FUNCTION_BLOCK R2 (* Basic Function Block Type *)
  (* Standard: 61499-2 *)
  (* Version 0.0, 10/11/2026, lizar, nxtControl GmBH, Template *)
  PACKAGE Main;
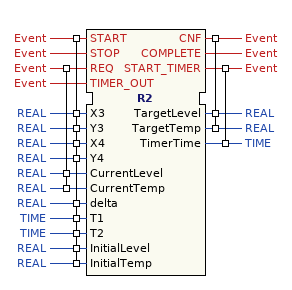
  EVENT_INPUT
    START WITH X3, Y3, X4, Y4, delta, T1, T2, InitialLevel, InitialTemp; (* Normal Execution Request *)
    STOP;
    REQ WITH CurrentLevel, CurrentTemp;
    TIMER_OUT;
  END_EVENT
  EVENT_OUTPUT
    CNF WITH TargetLevel, TargetTemp; (* Execution Confirmation *)
    COMPLETE;
    START_TIMER WITH TimerTime;
  END_EVENT
  VAR_INPUT
    X3 : REAL; (* Input event qualifier *)
    Y3 : REAL;
    X4 : REAL;
    Y4 : REAL;
    CurrentLevel : REAL;
    CurrentTemp : REAL;
    delta : REAL;
    T1 : TIME;
    T2 : TIME;
    InitialLevel : REAL;
    InitialTemp : REAL;
  END_VAR
  VAR_OUTPUT
    TargetLevel : REAL;
    TargetTemp : REAL;
    TimerTime : TIME;
  END_VAR
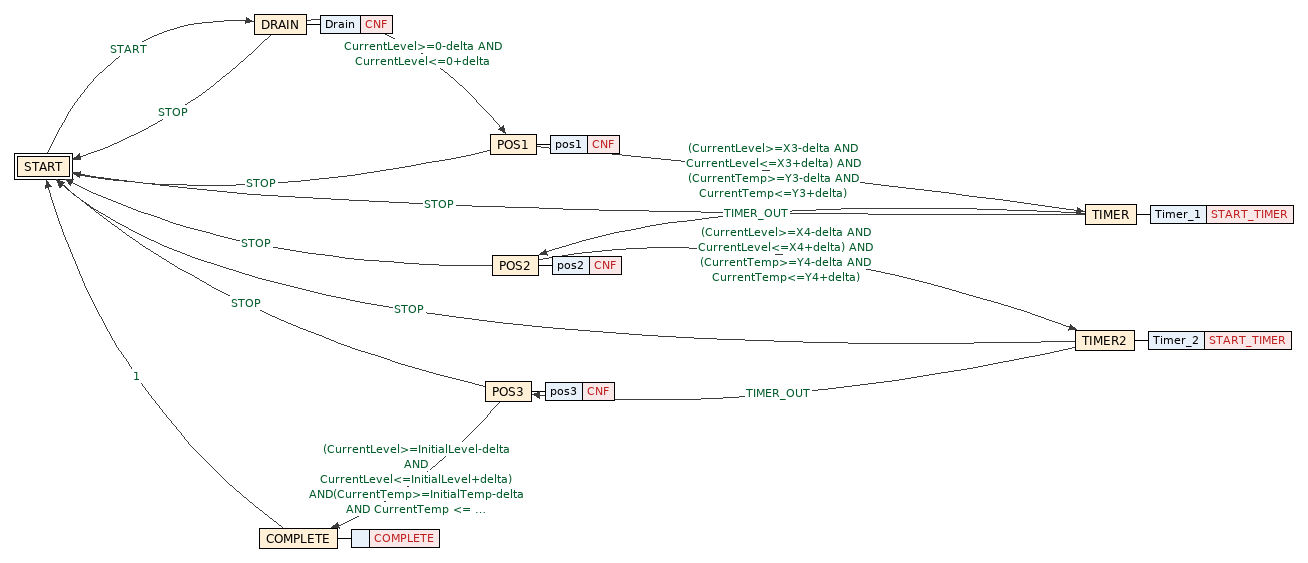
  EC_STATES
    START; (* Initial State *)
    DRAIN : Drain -> CNF;
    POS1 : pos1 -> CNF;
    POS2 : pos2 -> CNF;
    POS3 : pos3 -> CNF;
    COMPLETE : -> COMPLETE;
    TIMER : Timer_1 -> START_TIMER;
    TIMER2 : Timer_2 -> START_TIMER;
  END_STATES
  EC_TRANSITIONS
    START TO DRAIN := START;
    DRAIN TO POS1 := CurrentLevel>=0-delta AND CurrentLevel<=0+delta;
    POS3 TO COMPLETE := (CurrentLevel>=InitialLevel-delta AND CurrentLevel<=InitialLevel+delta) AND(CurrentTemp>=InitialTemp-delta AND CurrentTemp <= InitialTemp+delta);
    COMPLETE TO START := 1;
    DRAIN TO START := STOP;
    POS1 TO START := STOP;
    POS2 TO START := STOP;
    POS3 TO START := STOP;
    POS1 TO TIMER := (CurrentLevel>=X3-delta AND CurrentLevel<=X3+delta) AND (CurrentTemp>=Y3-delta AND CurrentTemp<=Y3+delta);
    TIMER TO POS2 := TIMER_OUT;
    POS2 TO TIMER2 := (CurrentLevel>=X4-delta AND CurrentLevel<=X4+delta) AND (CurrentTemp>=Y4-delta AND CurrentTemp<=Y4+delta);
    TIMER2 TO POS3 := TIMER_OUT;
    TIMER TO START := STOP;
    TIMER2 TO START := STOP;
  END_TRANSITIONS
  ALGORITHM Drain IN ST:
TargetLevel:= 0;
TargetTemp := 0;
  END_ALGORITHM
  ALGORITHM pos1 IN ST:
TargetLevel:= X3;
TargetTemp := Y3;
  END_ALGORITHM
  ALGORITHM pos2 IN ST:
TargetLevel:= X4;
TargetTemp := Y4;
  END_ALGORITHM
  ALGORITHM pos3 IN ST:
TargetLevel:= InitialLevel;
TargetTemp:= InitialTemp;
  END_ALGORITHM
  ALGORITHM Timer_1 IN ST:
TimerTime:= T1;
  END_ALGORITHM
  ALGORITHM Timer_2 IN ST:
TimerTime:= T2;
  END_ALGORITHM
END_FUNCTION_BLOCK
